Staubli VAL3: getDigIOSize.pgx

public program getDigIOSize(num& x_nSize)
  local num l_nSize
begin
  switch rs:sBusUsing
    case "MODBUS"
      l_nSize=size(_dInModbus)
    break
    case "PROFINET"
      l_nSize=size(_dInProfinet)
    break
    case "PROFIBUS"
      l_nSize=size(_dInProfibus)
    break
    case "ETHERCAT"
      l_nSize=size(_dInEtherCat)
    break
    case "ETHERNET"
      l_nSize=size(_dInEtherNet)
    break
  endSwitch
  x_nSize=l_nSize
end
